Staubli VAL3: deletePoint.pgx

public program deletePoint(string x_sKey, num x_nIndex, bool& x_bToSave)
  local bool l_bResult
begin
  l_bResult=userPageConfirm("是否删除点位："+toString("",x_nIndex))
  if l_bResult
    if x_nIndex==0 and size(trajTemp:tTrajItem[x_sKey].pPointItem)==1
      userPageAlert("数组元素不得为0")
    else
      delete(trajTemp:tTrajItem[x_sKey].pPointItem[x_nIndex])
      //trajTemp:libSave()
      x_bToSave=true
    endIf
  endIf

end
